// TIA Portal V20 export
// export: Created 2026-11-12T11:17:33.9569356Z, ExportSetting WithDefaults, DisplayName Totally Integrated Automation Portal, DisplayVersion V20, DisplayName TIA Portal Openness, DisplayVersion V20, DisplayName TIA Portal Teamcenter Gateway, DisplayVersion V20, DisplayName TIA Portal Version Control Interface, DisplayVersion V20, DisplayName STEP 7 Professional, DisplayVersion V20, DisplayName STEP 7 CFC, DisplayVersion V20, DisplayName STEP 7 Safety, DisplayVersion V20, DisplayName WinCC Basic/Comfort/Advanced, DisplayVersion V20, DisplayName SIMATIC Visualization Architect, DisplayVersion V20, DisplayName WinCC Professional, DisplayVersion V20, DisplayName SIMATIC Visualization Architect, DisplayVersion V20, DisplayName WinCC Unified, DisplayVersion V20, DisplayName SIMATIC Visualization Architect, DisplayVersion V20
TYPE "UDT_Estado"
// stored: IsFailsafeCompliant false
   STRUCT
      Modo_auto : Bool;   // Marca Modo
      Modo_manual : Bool;   // Marca Modo
      Ciclo_auto_activo : Bool;   // Marca Modo
      Ciclo_manual_activo : Bool;   // Marca Modo
      Emergencia : Bool;   // Marca Modo
      Rearme_requerido : Bool;   // Marca Modo
      Marcha_permitida : Bool;   // Marca Modo
      Condicion_arranque_auto : Bool;   // Marca Condiciones
      Condicion_arranque_manual : Bool;   // Marca Condiciones
      Estacion_cond_iniciales : Bool;   // Marca Condiciones
      Cinta_habilitada : Bool;   // Marca Condiciones
      Ciclo_manual_terminado : Bool;   // Marca Condiciones
      Rearme_requerido_gestion : Bool;   // Marca Condiciones
      Palet_en_posicion : Bool;   // Marca Cinta
      Palet_en_estacion : Bool;   // Marca Cinta
      Palet_evacuado : Bool;   // Marca Cinta
      Orden_evacuar : Bool;   // Marca Cinta
      Orden_leer : Bool;   // Marca RFID
      Orden_escribir : Bool;   // Marca RFID
      Rfid_lectura_ok : Bool;   // Marca RFID
      Rfid_escritura_ok : Bool;   // Marca RFID
      Rfid_error : Bool;   // Marca RFID
      Rfid_codigo_error : Byte;   // Marca RFID
      App_inicio : Bool;   // Marca App
      App_en_reposo : Bool;   // Marca App
      App_terminada : Bool;   // Marca App
      App_alarma : Bool;
   END_STRUCT;
END_TYPE
